(* IEC 61131-3 sources: esbmc-plc-benchmark-suite/benchmarks/manufacturing/st_comb_and, 1 file *)

(* ---- comb_and.st ---- *)
(* comb_and: three series contacts driving one coil.
   Structured Text rendering of ld_comb_and / g_comb_and.
   Y := A AND B AND C *)
PROGRAM drive
  VAR_INPUT
    A : BOOL;
    B : BOOL;
    C : BOOL;
  END_VAR
  VAR_OUTPUT
    Y : BOOL;
  END_VAR

  Y := A AND B AND C;
END_PROGRAM
